(* PLC project Vn_fn_concat, Beckhoff Automation GmbH TwinCAT PLC Control 3.5.13.21 *)
(* stored: creationDateTime 1970-01-01T00:00:00 *)

PROGRAM Vn_fn_concat

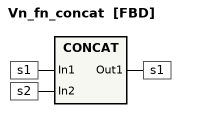
(* FBD diagram, written out as Structured Text *)
s1 := CONCAT(s1, s2);
END_PROGRAM
